TYPE TcoAbbRW_Outputs_v_8_2_x :
STRUCT
	Outputs AT %Q* : ARRAY[0..63] OF BYTE;
END_STRUCT
END_TYPE

(* stored: Version 1.1.0.1, ProductVersion 3.1.4024.12
   DUT TcoAbbRW_Outputs_v_8_2_x: Id {863ed5cc-fcd7-4b74-ae29-0b0a7103a64b} *)
